(* PLC project Deepseek3.project, CODESYS CODESYS V3.5 SP20 *)
(* stored: creationDateTime 2026-10-23T09:31:15.8733889, modificationDateTime 2026-10-23T09:31:05.9127754 *)

TYPE ST_Recipe : STRUCT
  sName : STRING(32);
  rMassSetpoint : REAL;  (* g *)
  tDripTime : TIME;  (* gotejamento *)
  tFillTimeout : TIME;  (* timeout de enchimento *)
END_STRUCT;
END_TYPE

TYPE E_DoseState : (IDLE := 0, LOCKING := 10, FILLING := 20, DRIPPING := 30, UNLOCKING := 40, DONE := 50, FAULT := 90);
END_TYPE

FUNCTION_BLOCK FB_FilterMovAvg
  VAR_INPUT
    rIn : REAL;  (* sinal de entrada *)
    nSamples : INT;  (* nº de amostras do buffer (1..100) *)
    xEnable : BOOL;  (* habilita atualização *)
  END_VAR
  VAR_OUTPUT
    rOut : REAL;  (* média móvel *)
  END_VAR
  VAR
    arBuffer : ARRAY[1..100] OF REAL;
    nIndex : INT := 1;
    nCount : INT;  (* amostras válidas no buffer *)
    i : INT;
    rSum : REAL;
    nEff : INT;
  END_VAR

                  (* Satura nº de amostras no limite do buffer *)
nEff := nSamples;
IF nEff < 1 THEN nEff := 1; END_IF
IF nEff > 100 THEN nEff := 100; END_IF

IF xEnable THEN
    (* Insere amostra (buffer circular) *)
    arBuffer[nIndex] := rIn;
    nIndex := nIndex + 1;
    IF nIndex > nEff THEN nIndex := 1; END_IF

    IF nCount < nEff THEN nCount := nCount + 1; END_IF

    (* Média móvel com laço FOR *)
    rSum := 0.0;
    FOR i := 1 TO nCount DO
        rSum := rSum + arBuffer[i];
    END_FOR
    IF nCount > 0 THEN
        rOut := rSum / INT_TO_REAL(nCount);
    END_IF
END_IF
                
END_FUNCTION_BLOCK

FUNCTION_BLOCK FB_ScaleAnalog
  VAR_INPUT
    nRaw : INT;
    rRawMin : REAL := 0.0;
    rRawMax : REAL := 27648.0;
    rEngMin : REAL;
    rEngMax : REAL;
  END_VAR
  VAR_OUTPUT
    rEng : REAL;
    xValid : BOOL;
  END_VAR

                  xValid := FALSE;
rEng   := rEngMin;   (* saída segura em falha *)

IF (rRawMax - rRawMin) <> 0.0 THEN
    rEng := rEngMin + (INT_TO_REAL(nRaw) - rRawMin) * (rEngMax - rEngMin) / (rRawMax - rRawMin);
END_IF

(* Validação simples de faixa bruta (com tolerância de under/overflow) *)
IF (nRaw >= -1000) AND (nRaw <= 28648) THEN
    xValid := TRUE;
END_IF
                
END_FUNCTION_BLOCK

FUNCTION_BLOCK FB_DosingLine
  VAR_INPUT
    xEnable : BOOL;  (* linha habilitada *)
    xMachineRun : BOOL;  (* ciclo automático ativo *)
    xBottlePresent : BOOL;  (* sensor de garrafa *)
    xCylExtended : BOOL;  (* fim de curso avançado *)
    xCylRetracted : BOOL;  (* fim de curso recolhido *)
    rMassActual : REAL;  (* massa atual (g) escalonada/filtrada *)
    rMassSetpoint : REAL;  (* massa alvo da receita (g) *)
    tDripTime : TIME;  (* tempo de gotejamento *)
    tFillTimeout : TIME;  (* tempo máximo de enchimento *)
    tCylMoveTimeout : TIME;  (* tempo máximo de movimento do cilindro *)
    xReset : BOOL;  (* reset de falhas *)
  END_VAR
  VAR_OUTPUT
    xLockCyl : BOOL;  (* comando trava garrafa *)
    xFillValve : BOOL;  (* comando válvula de enchimento *)
    xBusy : BOOL;  (* linha em ciclo *)
    xDone : BOOL;  (* ciclo desta linha concluído *)
    xBottleFilled : BOOL;  (* pulso: garrafa envasada *)
    xBottleRejected : BOOL;  (* pulso: garrafa rejeitada *)
    xFault : BOOL;  (* falha ativa da linha *)
    sFaultText : STRING(80);
    eState : E_DoseState;
  END_VAR
  VAR
    rtFillTO : TON;
    rtCylTO : TON;
    rtDrip : TON;
    rtPulse : TON;  (* alarga pulso de contagem *)
    xPrevDone : BOOL;
    xPrevFilled : BOOL;
    xPrevRejected : BOOL;
  END_VAR
  VAR CONSTANT
    tPulseWidth : TIME := TIME#100ms;  (* tempos internos de filtro de borda / pulso *)
  END_VAR

                  (* ------------------------------------------------------------- *)
(*  Pulsos de contagem: geração e auto-reset (largura fixa)      *)
(* ------------------------------------------------------------- *)
rtPulse(IN := xBottleFilled OR xBottleRejected, PT := tPulseWidth);
IF rtPulse.Q THEN
    xBottleFilled   := FALSE;
    xBottleRejected := FALSE;
END_IF

(* ------------------------------------------------------------- *)
(*  Reset global: limpa falhas e retorna à etapa IDLE            *)
(* ------------------------------------------------------------- *)
IF xReset THEN
    rtFillTO(IN := FALSE);
    rtCylTO (IN := FALSE);
    rtDrip  (IN := FALSE);
    xFault      := FALSE;
    sFaultText  := '';
    xLockCyl    := FALSE;
    xFillValve  := FALSE;
    eState      := E_DoseState.IDLE;
END_IF

(* ------------------------------------------------------------- *)
(*  Watchdog dos cilindros (tempo de movimento)                  *)
(* ------------------------------------------------------------- *)
rtCylTO(IN := (eState = E_DoseState.LOCKING) OR (eState = E_DoseState.UNLOCKING),
        PT := tCylMoveTimeout);
IF rtCylTO.Q AND NOT xFault THEN
    xFault     := TRUE;
    sFaultText := 'Timeout de movimento do cilindro';
    eState     := E_DoseState.FAULT;
END_IF

(* ------------------------------------------------------------- *)
(*  Watchdog de enchimento                                       *)
(* ------------------------------------------------------------- *)
rtFillTO(IN := (eState = E_DoseState.FILLING) OR (eState = E_DoseState.DRIPPING),
         PT := tFillTimeout);
IF rtFillTO.Q AND NOT xFault THEN
    xFault     := TRUE;
    sFaultText := 'Timeout de enchimento';
    eState     := E_DoseState.FAULT;
END_IF

(* ------------------------------------------------------------- *)
(*  Máquina de estados principal                                 *)
(* ------------------------------------------------------------- *)
CASE eState OF

    E_DoseState.IDLE:
        xLockCyl    := FALSE;
        xFillValve  := FALSE;
        xDone       := FALSE;
        xBusy       := FALSE;
        (* Só inicia se linha habilitada, ciclo ativo e garrafa presente *)
        IF xEnable AND xMachineRun AND xBottlePresent AND NOT xFault THEN
            xBusy  := TRUE;
            eState := E_DoseState.LOCKING;
        END_IF

    E_DoseState.LOCKING:
        xLockCyl := TRUE;
        IF xCylExtended THEN
            rtCylTO(IN := FALSE);
            eState := E_DoseState.FILLING;
        ELSIF NOT xBottlePresent THEN
            (* Garrafa removida durante a trava *)
            xFault     := TRUE;
            sFaultText := 'Garrafa removida durante o travamento';
            eState     := E_DoseState.FAULT;
        END_IF

    E_DoseState.FILLING:
        xLockCyl   := TRUE;
        xFillValve := TRUE;
        (* Garrafa removida durante o enchimento *)
        IF NOT xBottlePresent THEN
            xFillValve := FALSE;
            xFault     := TRUE;
            sFaultText := 'Garrafa removida durante o enchimento';
            eState     := E_DoseState.FAULT;
        ELSIF rMassActual >= rMassSetpoint THEN
            xFillValve := FALSE;
            rtDrip(IN := TRUE, PT := tDripTime);
            eState     := E_DoseState.DRIPPING;
        END_IF

    E_DoseState.DRIPPING:
        xLockCyl   := TRUE;
        xFillValve := FALSE;
        rtDrip(IN := TRUE, PT := tDripTime);
        IF rtDrip.Q THEN
            rtDrip(IN := FALSE);
            rtFillTO(IN := FALSE);
            eState := E_DoseState.UNLOCKING;
        END_IF

    E_DoseState.UNLOCKING:
        xLockCyl   := FALSE;
        xFillValve := FALSE;
        IF xCylRetracted THEN
            rtCylTO(IN := FALSE);
            xBottleFilled := TRUE;
            xDone         := TRUE;
            eState        := E_DoseState.DONE;
        END_IF

    E_DoseState.DONE:
        (* Mantém xDone até a esteira avançar; retorna a IDLE quando      *)
        (* a garrafa sai (sensor cai) ou o ciclo é reiniciado.            *)
        xLockCyl   := FALSE;
        xFillValve := FALSE;
        IF NOT xBottlePresent OR NOT xMachineRun THEN
            xDone  := FALSE;
            xBusy  := FALSE;
            eState := E_DoseState.IDLE;
        END_IF

    E_DoseState.FAULT:
        xLockCyl   := FALSE;
        xFillValve := FALSE;
        xFault     := TRUE;
        (* Linha permanece em falha até reset explícito *)
        IF NOT xBottlePresent THEN
            (* permite rejeição contabilizada pelo PRG_Main *)
        END_IF

END_CASE
                
END_FUNCTION_BLOCK

FUNCTION_BLOCK FB_TankLevel
  VAR_INPUT
    rLevelPct : REAL;  (* nível atual em % *)
    rLow : REAL := 30.0;  (* liga bomba *)
    rHigh : REAL := 80.0;  (* desliga bomba *)
    xMachineRun : BOOL;  (* se máquina parada, bomba pode parar *)
  END_VAR
  VAR_OUTPUT
    xPump : BOOL;
  END_VAR
  VAR
    xLatched : BOOL;
  END_VAR

                  (* Histerese: liga abaixo de rLow, desliga acima de rHigh *)
IF rLevelPct <= rLow THEN
    xLatched := TRUE;
ELSIF rLevelPct >= rHigh THEN
    xLatched := FALSE;
END_IF

(* Segurança: nível crítico baixo (<5%) força parada da bomba      *)
(* (evita cavitação; ajuste conforme o processo)                    *)
IF rLevelPct <= 5.0 THEN
    xLatched := FALSE;
END_IF

xPump := xLatched AND xMachineRun;
                
END_FUNCTION_BLOCK

FUNCTION_BLOCK FB_BottleCounter
  VAR_INPUT
    xFilledPulse : ARRAY[1..4] OF BOOL;  (* pulso por linha envasada *)
    xRejectedPulse : ARRAY[1..4] OF BOOL;  (* pulso por linha rejeitada *)
    xResetCounters : BOOL;
  END_VAR
  VAR_OUTPUT
    diFilled : DINT;
    diRejected : DINT;
  END_VAR
  VAR
    i : INT;
  END_VAR

                  IF xResetCounters THEN
    diFilled   := 0;
    diRejected := 0;
ELSE
    FOR i := 1 TO 4 DO
        IF xFilledPulse[i] THEN
            diFilled := diFilled + 1;
        END_IF
        IF xRejectedPulse[i] THEN
            diRejected := diRejected + 1;
        END_IF
    END_FOR
END_IF
                
END_FUNCTION_BLOCK

PROGRAM PRG_Main
  VAR
    fbScaleLoad : ARRAY[1..4] OF FB_ScaleAnalog;  (* Instâncias dos blocos funcionais *)
    fbAvgLoad : ARRAY[1..4] OF FB_FilterMovAvg;
    fbScaleTank : FB_ScaleAnalog;
    fbAvgTank : FB_FilterMovAvg;
    fbLines : ARRAY[1..4] OF FB_DosingLine;
    fbTank : FB_TankLevel;
    fbCounters : FB_BottleCounter;
    axBottleFilledPulse : ARRAY[1..4] OF BOOL;  (* Sinais derivados *)
    axBottleRejectPulse : ARRAY[1..4] OF BOOL;
    axLineFault : ARRAY[1..4] OF BOOL;
    axLineDone : ARRAY[1..4] OF BOOL;
    xAllLinesDone : BOOL;  (* Estado da esteira *)
    xAnyLineBusy : BOOL;
    xAnyLineFault : BOOL;
    rTankRawEng : REAL;  (* Escalonamento do nível do tanque *)
    stCurrentRecipe : ST_Recipe;  (* Receita corrente *)
    nRecipeSetpoint : INT;  (* Seleção de receita: só com máquina parada e nenhuma linha ativa *)
    i : INT;
    xAllLinesEnabled : BOOL;
  END_VAR

                  	(* ============================================================= *)
(*  1) EMERGÊNCIA E PORTA DE PROTEÇÃO — sobrepõem tudo           *)
(* ============================================================= *)
GVL_Main.xFaultGlobal := GVL_Main.xEmergStop OR NOT GVL_Main.xGuardDoor;

IF GVL_Main.xFaultGlobal THEN
    GVL_Main.xMachineRunning := FALSE;
    GVL_Main.xConveyorRun    := FALSE;
    FOR i := 1 TO 4 DO
        fbLines[i].xReset := TRUE;     (* força saída segura          *)
    END_FOR
    GVL_Main.xPumpTank := FALSE;
    GVL_Main.xLampGreen := FALSE;
    GVL_Main.xLampRed   := TRUE;
    GVL_Main.xHorn      := TRUE;
ELSE
    (* Reset normal: só com comando de reset e sem emergência *)
    IF GVL_Main.xResetPB THEN
        GVL_Main.xResetRequest := TRUE;
    END_IF
END_IF

(* Limpa pedido de reset após processamento *)
IF GVL_Main.xResetRequest AND NOT GVL_Main.xEmergStop AND GVL_Main.xGuardDoor THEN
    FOR i := 1 TO 4 DO
        fbLines[i].xReset := TRUE;
    END_FOR
    GVL_Main.xResetRequest := FALSE;
END_IF

(* ============================================================= *)
(*  2) SELEÇÃO DE RECEITA — apenas com máquina parada            *)
(* ============================================================= *)
xAllLinesEnabled := TRUE;
FOR i := 1 TO 4 DO
    IF NOT GVL_Main.axLineEnabled[i] THEN
        xAllLinesEnabled := FALSE;
    END_IF
END_FOR

nRecipeSetpoint := GVL_Main.nSelectedRecipe;
IF nRecipeSetpoint < 1 THEN nRecipeSetpoint := 1; END_IF
IF nRecipeSetpoint > 3 THEN nRecipeSetpoint := 3; END_IF

(* Receita só pode ser alterada se máquina parada e sem falhas     *)
(* (a atribuição direta já está protegida no HMI; aqui só copiamos) *)
stCurrentRecipe := GVL_Main.stRecipes[nRecipeSetpoint];

(* ============================================================= *)
(*  3) ESCALONAMENTO ANALÓGICO + MÉDIA MÓVEL                     *)
(* ============================================================= *)
FOR i := 1 TO 4 DO
    fbScaleLoad[i](
        nRaw    := GVL_Main.aiLoadCell[i],
        rRawMin := GVL_Main.rLoadCellRawMin,
        rRawMax := GVL_Main.rLoadCellRawMax,
        rEngMin := GVL_Main.rLoadCellEngMin,
        rEngMax := GVL_Main.rLoadCellEngMax
    );
    fbAvgLoad[i](
        rIn      := fbScaleLoad[i].rEng,
        nSamples := GVL_Main.nMovAvgSamples,
        xEnable  := NOT GVL_Main.xFaultGlobal
    );
    GVL_Main.arMassActual[i] := fbAvgLoad[i].rOut;
END_FOR

fbScaleTank(
    nRaw    := GVL_Main.aiTankLevel,
    rRawMin := GVL_Main.rTankRawMin,
    rRawMax := GVL_Main.rTankRawMax,
    rEngMin := GVL_Main.rTankEngMin,
    rEngMax := GVL_Main.rTankEngMax
);
fbAvgTank(
    rIn      := fbScaleTank.rEng,
    nSamples := GVL_Main.nMovAvgSamples,
    xEnable  := NOT GVL_Main.xFaultGlobal
);
GVL_Main.rTankLevelPct := fbAvgTank.rOut;

(* ============================================================= *)
(*  4) CONTROLE DE NÍVEL DO TANQUE (HISTERESE)                   *)
(* ============================================================= *)
fbTank(
    rLevelPct   := GVL_Main.rTankLevelPct,
    rLow        := GVL_Main.rTankLevelLow,
    rHigh       := GVL_Main.rTankLevelHigh,
    xMachineRun := GVL_Main.xMachineRunning
);
GVL_Main.xPumpTank := fbTank.xPump;

(* ============================================================= *)
(*  5) CICLO DE CADA LINHA DE ENCHIMENTO                         *)
(* ============================================================= *)
xAnyLineBusy  := FALSE;
xAnyLineFault := FALSE;
xAllLinesDone := TRUE;

FOR i := 1 TO 4 DO
    fbLines[i](
        xEnable         := GVL_Main.axLineEnabled[i] AND GVL_Main.xMachineRunning,
        xMachineRun     := GVL_Main.xMachineRunning,
        xBottlePresent  := GVL_Main.xBottlePresent[i],
        xCylExtended    := GVL_Main.xCylExtended[i],
        xCylRetracted   := GVL_Main.xCylRetracted[i],
        rMassActual     := GVL_Main.arMassActual[i],
        rMassSetpoint   := stCurrentRecipe.rMassSetpoint,
        tDripTime       := stCurrentRecipe.tDripTime,
        tFillTimeout    := stCurrentRecipe.tFillTimeout,
        tCylMoveTimeout := GVL_Main.tCylMoveTimeout,
        xReset          := FALSE
    );

    (* Saídas das linhas *)
    GVL_Main.xLockCyl[i]   := fbLines[i].xLockCyl;
    GVL_Main.xFillValve[i] := fbLines[i].xFillValve;

    (* Pulso de contagem e rejeição *)
    axBottleFilledPulse[i] := fbLines[i].xBottleFilled;
    (* Rejeição: falha ativa + garrafa presente = contabiliza descarte *)
    axBottleRejectPulse[i] := fbLines[i].xFault AND GVL_Main.xBottlePresent[i];

    axLineFault[i] := fbLines[i].xFault;
    axLineDone[i]  := fbLines[i].xDone;

    xAnyLineBusy  := xAnyLineBusy  OR fbLines[i].xBusy;
    xAnyLineFault := xAnyLineFault OR fbLines[i].xFault;

    (* Condição "linha concluída" considera linhas desabilitadas como prontas *)
    IF GVL_Main.axLineEnabled[i] THEN
        xAllLinesDone := xAllLinesDone AND fbLines[i].xDone;
    END_IF
END_FOR

(* ============================================================= *)
(*  6) FALHA GLOBAL AGREGADA + ALARMES                           *)
(* ============================================================= *)
IF xAnyLineFault OR GVL_Main.xFaultGlobal THEN
    GVL_Main.xLampRed   := TRUE;
    GVL_Main.xLampGreen := FALSE;
    GVL_Main.xHorn      := TRUE;
    GVL_Main.xMachineRunning := FALSE;
ELSE
    GVL_Main.xLampRed   := FALSE;
    GVL_Main.xHorn      := FALSE;
END_IF

(* ============================================================= *)
(*  7) COMANDO START/STOP                                        *)
(* ============================================================= *)
IF GVL_Main.xStartPB AND NOT GVL_Main.xFaultGlobal
   AND NOT xAnyLineFault AND GVL_Main.xGuardDoor
   AND NOT GVL_Main.xEmergStop THEN
    GVL_Main.xMachineRunning := TRUE;
END_IF

IF GVL_Main.xStopPB THEN
    GVL_Main.xMachineRunning := FALSE;
    GVL_Main.xConveyorRun    := FALSE;
END_IF

(* ============================================================= *)
(*  8) ESTEIRA: avança o próximo lote quando todas as linhas      *)
(*     habilitadas concluíram                                    *)
(* ============================================================= *)
IF GVL_Main.xMachineRunning AND NOT GVL_Main.xFaultGlobal
   AND NOT xAnyLineFault AND xAllLinesDone AND NOT xAnyLineBusy THEN
    (* Lote concluído: aciona esteira para próximo lote            *)
    IF GVL_Main.xConveyorPos THEN
        (* Ainda há lote posicionado — inicia avanço (retira lote) *)
        GVL_Main.xConveyorRun := TRUE;
    ELSE
        (* Novo lote posicionado — libera a esteira *)
        GVL_Main.xConveyorRun := FALSE;
    END_IF
END_IF

(* Se a esteira avançou e lote anterior saiu, reseta flags de DONE    *)
IF GVL_Main.xConveyorRun AND NOT GVL_Main.xConveyorPos THEN
    GVL_Main.xConveyorRun := FALSE;
END_IF

(* ============================================================= *)
(*  9) CONTADORES DE GARRAFAS                                    *)
(* ============================================================= *)
fbCounters(
    xFilledPulse   := axBottleFilledPulse,
    xRejectedPulse := axBottleRejectPulse,
    xResetCounters := FALSE
);
GVL_Main.diBottlesFilled   := fbCounters.diFilled;
GVL_Main.diBottlesRejected := fbCounters.diRejected;

(* ============================================================= *)
(* 10) SINALIZAÇÃO VERDE (máquina pronta / em ciclo)             *)
(* ============================================================= *)
IF GVL_Main.xMachineRunning AND NOT GVL_Main.xFaultGlobal AND NOT xAnyLineFault THEN
    GVL_Main.xLampGreen := TRUE;
END_IF
                
END_PROGRAM

CONFIGURATION Application
  RESOURCE Application ON PLC
    {attribute 'qualified_only'}
    VAR_GLOBAL  (* GVL_Main *)
      xEmergStop : BOOL;  (* 1 = emergência acionada (contato NF) *)
      xGuardDoor : BOOL;  (* 1 = porta de proteção FECHADA *)
      xStartPB : BOOL;  (* botão start *)
      xStopPB : BOOL;  (* botão stop *)
      xResetPB : BOOL;  (* botão reset de alarmes *)
      xBottlePresent : ARRAY[1..4] OF BOOL;  (* sensor de garrafa na linha *)
      xCylExtended : ARRAY[1..4] OF BOOL;  (* fim de curso cilindro avançado *)
      xCylRetracted : ARRAY[1..4] OF BOOL;  (* fim de curso cilindro recolhido *)
      xConveyorPos : BOOL;  (* lote posicionado (sensor de batente) *)
      aiLoadCell : ARRAY[1..4] OF INT;  (* célula de carga por linha 0..27648 *)
      aiTankLevel : INT;  (* nível do tanque 0..27648 *)
      xConveyorRun : BOOL;  (* aciona motor da esteira *)
      xLockCyl : ARRAY[1..4] OF BOOL;  (* trava garrafa (cilindro) *)
      xFillValve : ARRAY[1..4] OF BOOL;  (* válvula de enchimento *)
      xPumpTank : BOOL;  (* bomba de reposição do tanque pulmão *)
      xLampGreen : BOOL;
      xLampRed : BOOL;
      xHorn : BOOL;
      rLoadCellRawMin : REAL := 0.0;  (* valor bruto mínimo (INT) *)
      rLoadCellRawMax : REAL := 27648.0;  (* valor bruto máximo (INT) *)
      rLoadCellEngMin : REAL := 0.0;  (* 0 g *)
      rLoadCellEngMax : REAL := 5000.0;  (* 5000 g fundo de escala *)
      rTankRawMin : REAL := 0.0;
      rTankRawMax : REAL := 27648.0;
      rTankEngMin : REAL := 0.0;  (* 0 % *)
      rTankEngMax : REAL := 100.0;  (* 100 % *)
      nMovAvgSamples : INT := 10;  (* amostras da média móvel *)
      stRecipes : ARRAY[1..3] OF ST_Recipe := [(sName := 'R1 - 500g', rMassSetpoint := 500.0, tDripTime := TIME#300ms, tFillTimeout := TIME#15s0ms), (sName := 'R2 - 1000g', rMassSetpoint := 1000.0, tDripTime := TIME#400ms, tFillTimeout := TIME#20s0ms), (sName := 'R3 - 1500g', rMassSetpoint := 1500.0, tDripTime := TIME#500ms, tFillTimeout := TIME#25s0ms)];  (* ===================== RECEITAS =============================== [1..3] = receitas; [idx].rMassSetpoint em gramas *)
      nSelectedRecipe : INT := 1;  (* 1..3, alterável só com máquina parada *)
      axLineEnabled : ARRAY[1..4] OF BOOL := [TRUE, TRUE, TRUE, TRUE];  (* ===================== HABILITAÇÃO DE LINHAS ================== *)
      rTankLevelLow : REAL := 30.0;  (* % — liga bomba *)
      rTankLevelHigh : REAL := 80.0;  (* % — desliga bomba *)
      tCylMoveTimeout : TIME := TIME#3s0ms;  (* tempo máx. p/ cilindro mover *)
      xMachineRunning : BOOL;  (* ciclo automático habilitado *)
      xFaultGlobal : BOOL;  (* emergência ou porta aberta *)
      xResetRequest : BOOL;
      diBottlesFilled : DINT;  (* ===================== CONTADORES ============================= *)
      diBottlesRejected : DINT;
      arMassActual : ARRAY[1..4] OF REAL;  (* massa escalonada filtrada *)
      rTankLevelPct : REAL;
    END_VAR
    TASK MainTask(INTERVAL := T#20ms, PRIORITY := 1);
    PROGRAM PLC_PRG WITH MainTask : PLC_PRG;
  END_RESOURCE
END_CONFIGURATION
